Fanuc KAREL source: kx00025.compact.KL

PROGRAM KX00025
%COMMENT='Feature sample'
%STACKSIZE=65535
%PRIORITY=65535
%NOLOCKGROUP
VAR
I : INTEGER
J : INTEGER
B : BOOLEAN
F : FILE
S : STRING[80]
P : XYZWPR
BEGIN
I=1
END KX00025
